Fanuc KAREL source: ko00067.KL

-- PROVISIONAL review KL for V1013-1; original PC SHA256 a844cb2466df5f596a7c0082113837d4d7c8fa12b0d5a6651123cbff358bc4f3
-- Incomplete behavior may be omitted. Consult companion uncertainty JSON. Do not deploy.
PROGRAM KO00067
%NOLOCKGROUP
BEGIN
  -- UNRESOLVED_PC offsets 5-12; opcodes 9D,23
  -- UNRESOLVED_PC offsets 17-63; opcodes 27,22,1C,22,1C,22,31,7E,4A
  -- UNRESOLVED_PC offsets 68-72; opcodes 7F
END KO00067
